FUNCTION_BLOCK NOOP (* No-Op, auch bekannt als "No Operation" - reines Durchschleifen ohne internes FB *)
  (* Standard: 61131-3; Classification: standard boolean function; Description: Copyright (c) 2026 Meisterschulen am Ostbahnhof This program and the accompanying materials are made available under the terms of the Eclipse Public License 2.0 which is available at https://www.eclipse.org/legal/epl-2.0/ SPDX-License-Identifier: EPL-2.0 *)
  (* Version 1.1, 2026-10-11, Franz Höpfinger, Meisterschulen am Ostbahnhof, Copyright-Header, Classification und Remarks nachgezogen; Doku ergaenzt (kein internes FB, reiner Durchreicher) *)
  (* Version 1.0, 2026-05-05, franz, Meisterschulen am Ostbahnhof, initial API and implementation and/or initial documentation *)
  PACKAGE iec61131::booleanOperators;
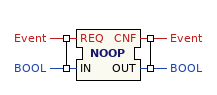
  EVENT_INPUT
    REQ WITH IN; (* Normal Execution Request *)
  END_EVENT
  EVENT_OUTPUT
    CNF WITH OUT; (* Execution Confirmation *)
  END_EVENT
  VAR_INPUT
    IN : BOOL; (* Input *)
  END_VAR
  VAR_OUTPUT
    OUT : BOOL; (* Output *)
  END_VAR
  EVENT_CONNECTIONS
    REQ TO CNF;
  END_CONNECTIONS
  DATA_CONNECTIONS
    IN TO OUT;
  END_CONNECTIONS
END_FUNCTION_BLOCK
